(* IEC 61131-3 sources: avi-aoi-management/scripts/ai-eval/ngau-nhien/kho/st-tt1-bo-phieu-2oo3/khung/src, 1 file *)

(* ---- BoPhieu2oo3.st ---- *)
FUNCTION_BLOCK BoPhieu2oo3
VAR_INPUT
    A : BOOL;
    B : BOOL;
    C : BOOL;
    RESET : BOOL;
END_VAR
VAR_OUTPUT
    Q : BOOL;
    LECH : BOOL;
    KENH_LECH : INT;
    DEM_LECH : DINT;
END_VAR
    (* TODO: cài đặt theo đề bài *)
    Q := FALSE;
END_FUNCTION_BLOCK
